(* IEC 61131-3 sources: codesys-to-s7/tests/corpus/C2S7-POU-FBINFC/neg, 1 file *)

(* ---- input.st ---- *)
FUNCTION_BLOCK FB_Case
VAR
    t : TON;
END_VAR
t(IN := TRUE, PT := T#1S);
END_FUNCTION_BLOCK
